{attribute 'qualified_only'}
{attribute 'strict'}
// Result of a manual focus re-home request (FB_FocusManualHome.Request).
TYPE E_FocusManualHome :
(
	Accepted := 0,
	NotAutomatic := 1,
	ManualUnlock := 2,
	AxisError := 3,
	NotCalibrated := 4,		// no longer returned (#138), kept for existing references
	Homing := 5,
	Moving := 6
);
END_TYPE

(* stored: Version 1.1.0.1, ProductVersion 3.1.4024.15
   DUT E_FocusManualHome: Id {a77ab252-d5df-4727-82c1-9790be8b2241} *)
